{attribute 'qualified_only'}
VAR_GLOBAL
	gvShutter1Up AT %Q* : BOOL;
END_VAR

(* stored: Version 1.1.0.1
   GVL GVL_Shutters: Id {7a0c2c86-f13b-43d1-9cdd-d1f7080b47ea} *)
